(*
    Tests of FB_AnalogInput16/32 (specs/analog-input).
*)
FUNCTION_BLOCK FB_AnalogInputTest EXTENDS TcUnit.FB_TestSuite
VAR
    AiNegative : MBIDivB.FB_AnalogInput16;
    AiElmNominal : MBIDivB.FB_AnalogInput32;
    AiElmPreset : MBIDivB.FB_AnalogInput32;
    AiZeroScale : MBIDivB.FB_AnalogInput16;
    AiConstant : MBIDivB.FB_AnalogInput16;
    AiReduced : MBIDivB.FB_AnalogInput16;
    AiSizeZero : MBIDivB.FB_AnalogInput16;
    AiOverrange : MBIDivB.FB_AnalogInput16;
    AiUnlinked : MBIDivB.FB_AnalogInput32;
    AiRestartStep : MBIDivB.FB_AnalogInput16;
    AiRestartSettings : MBIDivB.FB_AnalogInput32;
END_VAR


NegativeValue16Bit();
ElmNominalFullScale();
ElmExtendedPreset();
ZeroRawFullScaleRejected();
ConstantInputFiltered();
FilterSizeReducedRestarts();
FilterSizeZeroClampedToOne();
OverrangeSetAndCleared();
UnlinkedStatusBitsNoError();
RestartAfterStep();
RestartKeepsSettings();


METHOD PRIVATE ConstantInputFiltered
VAR
    Cycle : INT;
END_VAR

TEST('ConstantInputFiltered');

AiConstant.SetScale(RawFullScale := 1, ValueFullScale := 1.0);
AiConstant.Cfg.FilterSize := 10;
AiConstant.Raw := 2;
FOR Cycle := 1 TO 25 DO
    AiConstant();
END_FOR
AssertEquals_REAL(Expected := 2.0, Actual := AiConstant.Status.ValueFiltered, Delta := 1.0E-6, Message := 'ValueFiltered');

TEST_FINISHED();
END_METHOD


METHOD PRIVATE ElmExtendedPreset

TEST('ElmExtendedPreset');

AiElmPreset.SetScalePreset(Preset := MBIDivB.E_AiScalePreset.ELM3XXX_EXTENDED, NominalFullScale := 10.0);
AiElmPreset.Raw := 7812500;
AiElmPreset();
AssertEquals_REAL(Expected := 10.0, Actual := AiElmPreset.Status.Value, Delta := 1.0E-5, Message := 'nominal');
AiElmPreset.Raw := 8388607;
AiElmPreset();
AssertEquals_REAL(Expected := 10.737, Actual := AiElmPreset.Status.Value, Delta := 0.001, Message := 'technical full scale');

TEST_FINISHED();
END_METHOD


METHOD PRIVATE ElmNominalFullScale

TEST('ElmNominalFullScale');

AiElmNominal.SetScale(RawFullScale := 7812500, ValueFullScale := 10.0);
AiElmNominal.Raw := 7812500;
AiElmNominal();
AssertEquals_REAL(Expected := 10.0, Actual := AiElmNominal.Status.Value, Delta := 1.0E-5, Message := 'Value');
AssertEquals_DINT(Expected := 7812500, Actual := AiElmNominal.Status.RawFullScale, Message := 'RawFullScale');
AssertEquals_REAL(Expected := 10.0, Actual := AiElmNominal.Status.ValueFullScale, Delta := 1.0E-6, Message := 'ValueFullScale');

TEST_FINISHED();
END_METHOD


METHOD PRIVATE FilterSizeReducedRestarts
VAR
    Cycle : INT;
END_VAR

TEST('FilterSizeReducedRestarts');

AiReduced.SetScale(RawFullScale := 1, ValueFullScale := 1.0);
AiReduced.Cfg.FilterSize := 1000;
AiReduced.Raw := 3;
FOR Cycle := 1 TO 100 DO
    AiReduced();
END_FOR
AiReduced.Cfg.FilterSize := 10;
AiReduced.Raw := 1;
AiReduced();
AssertEquals_REAL(Expected := 1.0, Actual := AiReduced.Status.ValueFiltered, Delta := 1.0E-6, Message := 'no contribution from older samples');

TEST_FINISHED();
END_METHOD


METHOD PRIVATE FilterSizeZeroClampedToOne

TEST('FilterSizeZeroClampedToOne');

AiSizeZero.SetScale(RawFullScale := 1, ValueFullScale := 1.0);
AiSizeZero.Cfg.FilterSize := 0;
AiSizeZero.Raw := 4;
AiSizeZero();
AssertEquals_DINT(Expected := 1, Actual := AiSizeZero.Cfg.FilterSize, Message := 'FilterSize written back');
AssertEquals_REAL(Expected := 4.0, Actual := AiSizeZero.Status.ValueFiltered, Delta := 1.0E-6, Message := 'ValueFiltered');

TEST_FINISHED();
END_METHOD


METHOD PRIVATE NegativeValue16Bit

TEST('NegativeValue16Bit');

AiNegative.SetScalePreset(Preset := MBIDivB.E_AiScalePreset.EL31XX_LEGACY, NominalFullScale := 10.0);
AiNegative.Raw := -16384;
AiNegative();
AssertEquals_REAL(Expected := -5.0, Actual := AiNegative.Status.Value, Delta := 0.001, Message := 'Value');
AssertEquals_DINT(Expected := -16384, Actual := AiNegative.Status.Raw, Message := 'Raw');

TEST_FINISHED();
END_METHOD


METHOD PRIVATE OverrangeSetAndCleared

TEST('OverrangeSetAndCleared');

AiOverrange.Overrange := TRUE;
AiOverrange();
AssertTrue(Condition := AiOverrange.Status.Error, Message := 'Error while set');
AssertTrue(Condition := FIND(AiOverrange.Status.ErrorText, 'overrange') > 0, Message := 'ErrorText mentions overrange');
AiOverrange.Overrange := FALSE;
AiOverrange();
AssertFalse(Condition := AiOverrange.Status.Error, Message := 'Error cleared');
AssertEquals_STRING(Expected := '', Actual := AiOverrange.Status.ErrorText, Message := 'ErrorText cleared');

TEST_FINISHED();
END_METHOD


METHOD PRIVATE RestartAfterStep
VAR
    Cycle : INT;
    Wrong : INT;
END_VAR

TEST('RestartAfterStep');

AiRestartStep.SetScale(RawFullScale := 1000, ValueFullScale := 1.0);
AiRestartStep.Cfg.FilterSize := 10;
AiRestartStep.Raw := 1000;
FOR Cycle := 1 TO 15 DO
    AiRestartStep();
END_FOR
AiRestartStep.RestartFilter();
AiRestartStep.Raw := 3000;
FOR Cycle := 1 TO 12 DO
    AiRestartStep();
    IF ABS(AiRestartStep.Status.ValueFiltered - 3.0) > 1.0E-6 THEN
        Wrong := Wrong + 1;
    END_IF
END_FOR
AssertEquals_INT(Expected := 0, Actual := Wrong, Message := 'calls with ValueFiltered <> 3.0 V after the restart');

TEST_FINISHED();
END_METHOD


METHOD PRIVATE RestartKeepsSettings

TEST('RestartKeepsSettings');

AiRestartSettings.SetScale(RawFullScale := 7812500, ValueFullScale := 10.0);
AiRestartSettings.Cfg.FilterSize := 20;
AiRestartSettings.Raw := 3906250;
AiRestartSettings();
AiRestartSettings.RestartFilter();
AiRestartSettings();
AssertEquals_DINT(Expected := 20, Actual := AiRestartSettings.Cfg.FilterSize, Message := 'FilterSize');
AssertEquals_DINT(Expected := 7812500, Actual := AiRestartSettings.Status.RawFullScale, Message := 'RawFullScale');
AssertEquals_REAL(Expected := 10.0, Actual := AiRestartSettings.Status.ValueFullScale, Delta := 1.0E-6, Message := 'ValueFullScale');
AssertEquals_REAL(Expected := 5.0, Actual := AiRestartSettings.Status.Value, Delta := 1.0E-5, Message := 'Value');

TEST_FINISHED();
END_METHOD


METHOD PRIVATE UnlinkedStatusBitsNoError

TEST('UnlinkedStatusBitsNoError');

AiUnlinked.Raw := 1000;
AiUnlinked();
AssertFalse(Condition := AiUnlinked.Status.Error, Message := 'Error');

TEST_FINISHED();
END_METHOD


METHOD PRIVATE ZeroRawFullScaleRejected
VAR
    Accepted : BOOL;
END_VAR

TEST('ZeroRawFullScaleRejected');

AiZeroScale.SetScale(RawFullScale := 32767, ValueFullScale := 10.0);
Accepted := AiZeroScale.SetScale(RawFullScale := 0, ValueFullScale := 5.0);
AiZeroScale.Raw := 16384;
AiZeroScale();
AssertFalse(Condition := Accepted, Message := 'SetScale must return FALSE');
AssertTrue(Condition := AiZeroScale.Status.Error, Message := 'Error');
AssertTrue(Condition := FIND(AiZeroScale.Status.ErrorText, 'RawFullScale') > 0, Message := 'ErrorText names RawFullScale');
AssertEquals_REAL(Expected := 5.0, Actual := AiZeroScale.Status.Value, Delta := 0.001, Message := 'previous scaling kept');

TEST_FINISHED();
END_METHOD

END_FUNCTION_BLOCK

(* stored: Version 1.1.0.1
   POU FB_AnalogInputTest: Id {5e6b4b2d-4371-4b29-b5d9-ec526945e7b8}, SpecialFunc None
   Method ConstantInputFiltered: Id {faae7e18-d223-4327-8ed7-bf86f08b6b7b}
   Method ElmExtendedPreset: Id {a093f940-8ef6-4efb-bd02-eb0bfaa95578}
   Method ElmNominalFullScale: Id {5aa880d2-43fe-4984-9814-6bfecdfc0b07}
   Method FilterSizeReducedRestarts: Id {9e393518-3ba6-4299-b581-cff858c7566c}
   Method FilterSizeZeroClampedToOne: Id {3f728ffe-d033-49c7-9656-490115839e3a}
   Method NegativeValue16Bit: Id {1477b943-c372-476e-b432-8f8c9dd0c34b}
   Method OverrangeSetAndCleared: Id {d71aeace-9d3e-424c-aea7-ea346418a1c4}
   Method RestartAfterStep: Id {ed0fd9de-e843-4d79-a4b9-df14db3fe521}
   Method RestartKeepsSettings: Id {ffbeb672-e086-4675-9341-5f0d5534fa92}
   Method UnlinkedStatusBitsNoError: Id {b38776f0-790e-4f83-9a9f-b384b076d963}
   Method ZeroRawFullScaleRejected: Id {42d319a6-c1e0-427f-88c8-41bd2d9ed738} *)
